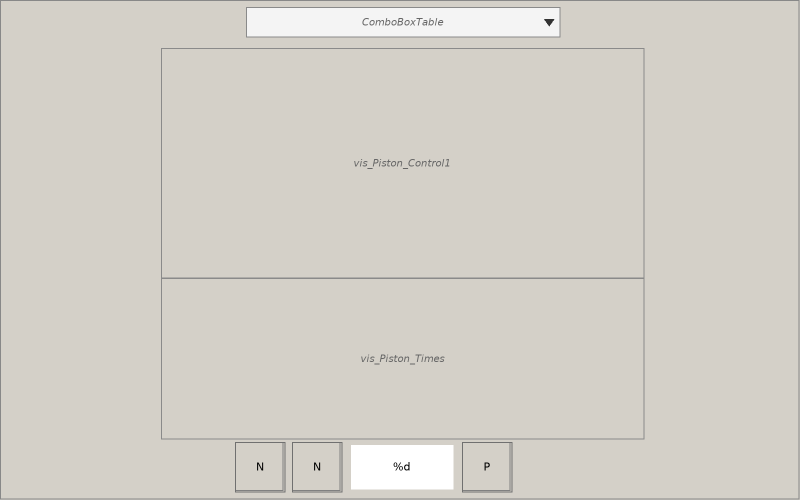
VISUALIZATION vis_Piston_Select  // 800x500
    Frame (161,48 483x230)
        shows vis_Piston_Control1(stPis := stPis[iPis_sel])
    Frame (161,278 483x161)
        shows vis_Piston_Times(stPis := stPis[iPis_sel])
    Button (292,442 50x50), "N"
        tap prg_Piston.bPis_Next_N
    Button (462,442 50x50), "P"
        tap prg_Piston.bPis_Next_P
    Textfield (350,444 104x46), "%d", text variable: iPis_sel
    ComboBoxTable (246,7 314x30), variable: iPis_sel, data array: g_Piston.arPisName
        p3854506369: g_Piston.arPisName[INDEX].Num
        p1892666644: g_Piston.arPisName[INDEX].Description
    Button (235,442 50x50), "N"
        tap prg_Piston.bPis_Next_N
END_VISUALIZATION

(* stored: Version 1.1.0.1, ProductVersion 3.1.4024.12
   Visu vis_Piston_Select: Id {0a1b4940-e1fb-4049-b08d-892a3c8e3439} *)
